FUNCTION FC 1 : VOID
BEGIN
NETWORK
      L S5T#1S5MS
END_FUNCTION
